// TIA Portal V21 export
// export: Created 2026-11-21T13:26:59.0904116Z, ExportSetting WithDefaults, DisplayName Totally Integrated Automation Portal, DisplayVersion V21, DisplayName STEP 7 Professional, DisplayVersion V21, DisplayName STEP 7 Safety, DisplayVersion V21, DisplayName Tech WebApplication, DisplayVersion V21, DisplayName WinCC Basic/Comfort/Advanced, DisplayVersion V21, DisplayName WinCC Unified, DisplayVersion V21
VAR_GLOBAL   // PLC tag table "Signals"
   levelSensor AT %IW10 : Int;   // Füllstandsensor / Level sensor / Capteur de niveau
   pumpOn AT %Q4.0 : Bool;   // Pumpe ein / Pump on / Pompe en marche
   spare AT %Q4.1 : Bool;   // Spare output
END_VAR
